// TIA Portal V21 export
// export: Created 2026-11-08T21:21:56.8202802Z, ExportSetting WithDefaults, DisplayName Totally Integrated Automation Portal, DisplayVersion V21 Update 3, DisplayName STEP 7 Professional, DisplayVersion V21 Update 3, DisplayName STEP 7 Safety, DisplayVersion V21, DisplayName Tech WebApplication, DisplayVersion V21, DisplayName WinCC Basic/Comfort/Advanced, DisplayVersion V21 Update 3, DisplayName WinCC Unified, DisplayVersion V21 Update 3
FUNCTION_BLOCK "FB_Graph"   // FB74, GRAPH
VERSION : 0.1
// stored: AcknowledgeErrorsRequired true, AutoNumber true, GraphVersion 6.0, InitialValuesAcquisition false, IsIECCheckEnabled false, LanguageInNetworks LAD, LockOperatingMode false, PermanentILProcessingInMANMode false, SetENOAutomatically false, SkipSteps false, UDAEnableTagReadback false, WithAlarmHandling true
   // inherited from GRAPH_BASE
   VAR
      OFF_SQ_BASE : Bool;
   END_VAR
   VAR_INPUT
      OFF_SQ : Bool := false;   // Turn sequence off
      INIT_SQ : Bool := false;   // Set sequence to initial state
      ACK_EF : Bool := false;   // Acknowledge all errors and faults
      go : Bool;
      "a" : Bool;
      "b" : Bool;
      sv : Bool;
   END_VAR
   VAR_OUTPUT
      q1 : Bool;
      q2 : Bool;
      q3 : Bool;
   END_VAR
BEGIN
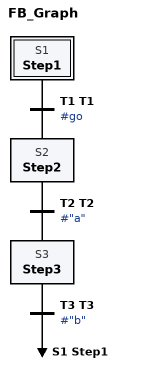
   // sequencer 1
   INITIAL_STEP Step1:   // S1, max time T#10S, warning time T#7S
      supervision V := #sv;
   END_STEP
   TRANSITION T1 FROM Step1 TO Step2   // T1
      := #go;
   END_TRANSITION
   STEP Step2:   // S2, max time T#10S, warning time T#7S
      supervision V := #sv;
   END_STEP
   TRANSITION T2 FROM Step2 TO Step3   // T2
      := #"a";
   END_TRANSITION
   STEP Step3:   // S3, max time T#10S, warning time T#7S
      supervision V := #sv;
   END_STEP
   TRANSITION T3 FROM Step3 TO Step1   // T3, jump
      := #"b";
   END_TRANSITION
END_FUNCTION_BLOCK
